(* IEC 61131-3 sources: sis-interlock-demo/tests/POUs/TruthTables/FB_VoteTableFbSmall_Test, 18 files *)

(* ---- Fb1oo1DAAIMatchesModel.method.decl.st ---- *)
// AUTO-GENERATED by tools_project/gen_voting_tests.py — не редактировать: правьте генератор или модель
//   tools_project/vote_model.py и запустите python tools_project/gen_voting_tests.py
// FB_Voting, схема 1oo1, политика DA, вход AI: все 8 сочетаний
// (требование × достоверность × запрос байпаса по каналу — для FB_Voting); ожидаемые значения —
// эталонная модель tools_project/vote_model.py. Один AssertEquals_BYTE на строку.
METHOD PRIVATE Fb1oo1DAAIMatchesModel
VAR
    fbRig : FB_VoteTableRig;   // стенд таблиц (новый экземпляр на тест)
    bRes  : BYTE;              // код результата строки
END_VAR

(* ---- Fb1oo1DADIMatchesModel.method.decl.st ---- *)
// AUTO-GENERATED by tools_project/gen_voting_tests.py — не редактировать: правьте генератор или модель
//   tools_project/vote_model.py и запустите python tools_project/gen_voting_tests.py
// FB_Voting, схема 1oo1, политика DA, вход DI: все 8 сочетаний
// (требование × достоверность × запрос байпаса по каналу — для FB_Voting); ожидаемые значения —
// эталонная модель tools_project/vote_model.py. Один AssertEquals_BYTE на строку.
METHOD PRIVATE Fb1oo1DADIMatchesModel
VAR
    fbRig : FB_VoteTableRig;   // стенд таблиц (новый экземпляр на тест)
    bRes  : BYTE;              // код результата строки
END_VAR

(* ---- Fb1oo1DSAIMatchesModel.method.decl.st ---- *)
// AUTO-GENERATED by tools_project/gen_voting_tests.py — не редактировать: правьте генератор или модель
//   tools_project/vote_model.py и запустите python tools_project/gen_voting_tests.py
// FB_Voting, схема 1oo1, политика DS, вход AI: все 8 сочетаний
// (требование × достоверность × запрос байпаса по каналу — для FB_Voting); ожидаемые значения —
// эталонная модель tools_project/vote_model.py. Один AssertEquals_BYTE на строку.
METHOD PRIVATE Fb1oo1DSAIMatchesModel
VAR
    fbRig : FB_VoteTableRig;   // стенд таблиц (новый экземпляр на тест)
    bRes  : BYTE;              // код результата строки
END_VAR

(* ---- Fb1oo1DSDIMatchesModel.method.decl.st ---- *)
// AUTO-GENERATED by tools_project/gen_voting_tests.py — не редактировать: правьте генератор или модель
//   tools_project/vote_model.py и запустите python tools_project/gen_voting_tests.py
// FB_Voting, схема 1oo1, политика DS, вход DI: все 8 сочетаний
// (требование × достоверность × запрос байпаса по каналу — для FB_Voting); ожидаемые значения —
// эталонная модель tools_project/vote_model.py. Один AssertEquals_BYTE на строку.
METHOD PRIVATE Fb1oo1DSDIMatchesModel
VAR
    fbRig : FB_VoteTableRig;   // стенд таблиц (новый экземпляр на тест)
    bRes  : BYTE;              // код результата строки
END_VAR

(* ---- Fb1oo1VTAIMatchesModel.method.decl.st ---- *)
// AUTO-GENERATED by tools_project/gen_voting_tests.py — не редактировать: правьте генератор или модель
//   tools_project/vote_model.py и запустите python tools_project/gen_voting_tests.py
// FB_Voting, схема 1oo1, политика VT, вход AI: все 8 сочетаний
// (требование × достоверность × запрос байпаса по каналу — для FB_Voting); ожидаемые значения —
// эталонная модель tools_project/vote_model.py. Один AssertEquals_BYTE на строку.
METHOD PRIVATE Fb1oo1VTAIMatchesModel
VAR
    fbRig : FB_VoteTableRig;   // стенд таблиц (новый экземпляр на тест)
    bRes  : BYTE;              // код результата строки
END_VAR

(* ---- Fb1oo1VTDIMatchesModel.method.decl.st ---- *)
// AUTO-GENERATED by tools_project/gen_voting_tests.py — не редактировать: правьте генератор или модель
//   tools_project/vote_model.py и запустите python tools_project/gen_voting_tests.py
// FB_Voting, схема 1oo1, политика VT, вход DI: все 8 сочетаний
// (требование × достоверность × запрос байпаса по каналу — для FB_Voting); ожидаемые значения —
// эталонная модель tools_project/vote_model.py. Один AssertEquals_BYTE на строку.
METHOD PRIVATE Fb1oo1VTDIMatchesModel
VAR
    fbRig : FB_VoteTableRig;   // стенд таблиц (новый экземпляр на тест)
    bRes  : BYTE;              // код результата строки
END_VAR

(* ---- Fb1oo2DAAIMatchesModel.method.decl.st ---- *)
// AUTO-GENERATED by tools_project/gen_voting_tests.py — не редактировать: правьте генератор или модель
//   tools_project/vote_model.py и запустите python tools_project/gen_voting_tests.py
// FB_Voting, схема 1oo2, политика DA, вход AI: все 64 сочетаний
// (требование × достоверность × запрос байпаса по каналу — для FB_Voting); ожидаемые значения —
// эталонная модель tools_project/vote_model.py. Один AssertEquals_BYTE на строку.
METHOD PRIVATE Fb1oo2DAAIMatchesModel
VAR
    fbRig : FB_VoteTableRig;   // стенд таблиц (новый экземпляр на тест)
    bRes  : BYTE;              // код результата строки
END_VAR

(* ---- Fb1oo2DADIMatchesModel.method.decl.st ---- *)
// AUTO-GENERATED by tools_project/gen_voting_tests.py — не редактировать: правьте генератор или модель
//   tools_project/vote_model.py и запустите python tools_project/gen_voting_tests.py
// FB_Voting, схема 1oo2, политика DA, вход DI: все 64 сочетаний
// (требование × достоверность × запрос байпаса по каналу — для FB_Voting); ожидаемые значения —
// эталонная модель tools_project/vote_model.py. Один AssertEquals_BYTE на строку.
METHOD PRIVATE Fb1oo2DADIMatchesModel
VAR
    fbRig : FB_VoteTableRig;   // стенд таблиц (новый экземпляр на тест)
    bRes  : BYTE;              // код результата строки
END_VAR

(* ---- Fb1oo2DSAIMatchesModel.method.decl.st ---- *)
// AUTO-GENERATED by tools_project/gen_voting_tests.py — не редактировать: правьте генератор или модель
//   tools_project/vote_model.py и запустите python tools_project/gen_voting_tests.py
// FB_Voting, схема 1oo2, политика DS, вход AI: все 64 сочетаний
// (требование × достоверность × запрос байпаса по каналу — для FB_Voting); ожидаемые значения —
// эталонная модель tools_project/vote_model.py. Один AssertEquals_BYTE на строку.
METHOD PRIVATE Fb1oo2DSAIMatchesModel
VAR
    fbRig : FB_VoteTableRig;   // стенд таблиц (новый экземпляр на тест)
    bRes  : BYTE;              // код результата строки
END_VAR

(* ---- Fb1oo2DSDIMatchesModel.method.decl.st ---- *)
// AUTO-GENERATED by tools_project/gen_voting_tests.py — не редактировать: правьте генератор или модель
//   tools_project/vote_model.py и запустите python tools_project/gen_voting_tests.py
// FB_Voting, схема 1oo2, политика DS, вход DI: все 64 сочетаний
// (требование × достоверность × запрос байпаса по каналу — для FB_Voting); ожидаемые значения —
// эталонная модель tools_project/vote_model.py. Один AssertEquals_BYTE на строку.
METHOD PRIVATE Fb1oo2DSDIMatchesModel
VAR
    fbRig : FB_VoteTableRig;   // стенд таблиц (новый экземпляр на тест)
    bRes  : BYTE;              // код результата строки
END_VAR

(* ---- Fb1oo2VTAIMatchesModel.method.decl.st ---- *)
// AUTO-GENERATED by tools_project/gen_voting_tests.py — не редактировать: правьте генератор или модель
//   tools_project/vote_model.py и запустите python tools_project/gen_voting_tests.py
// FB_Voting, схема 1oo2, политика VT, вход AI: все 64 сочетаний
// (требование × достоверность × запрос байпаса по каналу — для FB_Voting); ожидаемые значения —
// эталонная модель tools_project/vote_model.py. Один AssertEquals_BYTE на строку.
METHOD PRIVATE Fb1oo2VTAIMatchesModel
VAR
    fbRig : FB_VoteTableRig;   // стенд таблиц (новый экземпляр на тест)
    bRes  : BYTE;              // код результата строки
END_VAR

(* ---- Fb1oo2VTDIMatchesModel.method.decl.st ---- *)
// AUTO-GENERATED by tools_project/gen_voting_tests.py — не редактировать: правьте генератор или модель
//   tools_project/vote_model.py и запустите python tools_project/gen_voting_tests.py
// FB_Voting, схема 1oo2, политика VT, вход DI: все 64 сочетаний
// (требование × достоверность × запрос байпаса по каналу — для FB_Voting); ожидаемые значения —
// эталонная модель tools_project/vote_model.py. Один AssertEquals_BYTE на строку.
METHOD PRIVATE Fb1oo2VTDIMatchesModel
VAR
    fbRig : FB_VoteTableRig;   // стенд таблиц (новый экземпляр на тест)
    bRes  : BYTE;              // код результата строки
END_VAR

(* ---- Fb2oo2DAAIMatchesModel.method.decl.st ---- *)
// AUTO-GENERATED by tools_project/gen_voting_tests.py — не редактировать: правьте генератор или модель
//   tools_project/vote_model.py и запустите python tools_project/gen_voting_tests.py
// FB_Voting, схема 2oo2, политика DA, вход AI: все 64 сочетаний
// (требование × достоверность × запрос байпаса по каналу — для FB_Voting); ожидаемые значения —
// эталонная модель tools_project/vote_model.py. Один AssertEquals_BYTE на строку.
METHOD PRIVATE Fb2oo2DAAIMatchesModel
VAR
    fbRig : FB_VoteTableRig;   // стенд таблиц (новый экземпляр на тест)
    bRes  : BYTE;              // код результата строки
END_VAR

(* ---- Fb2oo2DADIMatchesModel.method.decl.st ---- *)
// AUTO-GENERATED by tools_project/gen_voting_tests.py — не редактировать: правьте генератор или модель
//   tools_project/vote_model.py и запустите python tools_project/gen_voting_tests.py
// FB_Voting, схема 2oo2, политика DA, вход DI: все 64 сочетаний
// (требование × достоверность × запрос байпаса по каналу — для FB_Voting); ожидаемые значения —
// эталонная модель tools_project/vote_model.py. Один AssertEquals_BYTE на строку.
METHOD PRIVATE Fb2oo2DADIMatchesModel
VAR
    fbRig : FB_VoteTableRig;   // стенд таблиц (новый экземпляр на тест)
    bRes  : BYTE;              // код результата строки
END_VAR

(* ---- Fb2oo2DSAIMatchesModel.method.decl.st ---- *)
// AUTO-GENERATED by tools_project/gen_voting_tests.py — не редактировать: правьте генератор или модель
//   tools_project/vote_model.py и запустите python tools_project/gen_voting_tests.py
// FB_Voting, схема 2oo2, политика DS, вход AI: все 64 сочетаний
// (требование × достоверность × запрос байпаса по каналу — для FB_Voting); ожидаемые значения —
// эталонная модель tools_project/vote_model.py. Один AssertEquals_BYTE на строку.
METHOD PRIVATE Fb2oo2DSAIMatchesModel
VAR
    fbRig : FB_VoteTableRig;   // стенд таблиц (новый экземпляр на тест)
    bRes  : BYTE;              // код результата строки
END_VAR

(* ---- Fb2oo2DSDIMatchesModel.method.decl.st ---- *)
// AUTO-GENERATED by tools_project/gen_voting_tests.py — не редактировать: правьте генератор или модель
//   tools_project/vote_model.py и запустите python tools_project/gen_voting_tests.py
// FB_Voting, схема 2oo2, политика DS, вход DI: все 64 сочетаний
// (требование × достоверность × запрос байпаса по каналу — для FB_Voting); ожидаемые значения —
// эталонная модель tools_project/vote_model.py. Один AssertEquals_BYTE на строку.
METHOD PRIVATE Fb2oo2DSDIMatchesModel
VAR
    fbRig : FB_VoteTableRig;   // стенд таблиц (новый экземпляр на тест)
    bRes  : BYTE;              // код результата строки
END_VAR

(* ---- Fb2oo2VTAIMatchesModel.method.decl.st ---- *)
// AUTO-GENERATED by tools_project/gen_voting_tests.py — не редактировать: правьте генератор или модель
//   tools_project/vote_model.py и запустите python tools_project/gen_voting_tests.py
// FB_Voting, схема 2oo2, политика VT, вход AI: все 64 сочетаний
// (требование × достоверность × запрос байпаса по каналу — для FB_Voting); ожидаемые значения —
// эталонная модель tools_project/vote_model.py. Один AssertEquals_BYTE на строку.
METHOD PRIVATE Fb2oo2VTAIMatchesModel
VAR
    fbRig : FB_VoteTableRig;   // стенд таблиц (новый экземпляр на тест)
    bRes  : BYTE;              // код результата строки
END_VAR

(* ---- Fb2oo2VTDIMatchesModel.method.decl.st ---- *)
// AUTO-GENERATED by tools_project/gen_voting_tests.py — не редактировать: правьте генератор или модель
//   tools_project/vote_model.py и запустите python tools_project/gen_voting_tests.py
// FB_Voting, схема 2oo2, политика VT, вход DI: все 64 сочетаний
// (требование × достоверность × запрос байпаса по каналу — для FB_Voting); ожидаемые значения —
// эталонная модель tools_project/vote_model.py. Один AssertEquals_BYTE на строку.
METHOD PRIVATE Fb2oo2VTDIMatchesModel
VAR
    fbRig : FB_VoteTableRig;   // стенд таблиц (новый экземпляр на тест)
    bRes  : BYTE;              // код результата строки
END_VAR
